// TIA Portal V20 export
Screen "ALARM_HISTORY"  1276x673
  ScreenItem "Title_ScreenOverview_X390_Y2" at 390,2 size 510x57  Type=HmiTextBox
  ScreenItem "Alarm_History_Legend" at 1180,2 size 90x60  Type=HmiButton
  ScreenItem "permanentareaborderrectangle" at 0,0 size 0x0  Type=HmiRectangle
  ScreenItem "Line_Header_X0_Y64_1" at 0,64 size 1280x0  Type=HmiLine
  ScreenItem "Button_Back" at 2,2 size 90x60  Type=HmiButton
  ScreenItem "Button_Language" at 97,2 size 90x60  Type=HmiButton
  ScreenItem "报警控件_1" at 0,66 size 1280x602  Type=HmiAlarmControl
  ScreenItem "Line_Header_X0_Y64_2" at 0,64 size 1276x0  Type=HmiLine
  ScreenItem "txtClearHistory" at 193,2 size 90x60  Type=HmiTextBox
